// Mitsubishi GX Works2 project: 적산타이머   PLC: Q02/Q02H

PROGRAM MAIN
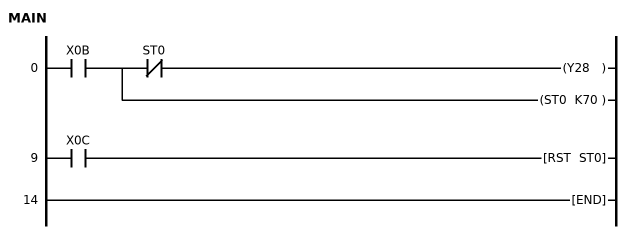
0     LD      X0B
      MPS
      ANI     ST0
      OUT     Y28
      MPP
      OUT     ST0 K70
9     LD      X0C
      RST     ST0
14    END
END_PROGRAM
